(* IEC 61131-3 sources: SortJet_MasterSPS_Aufbau.fbsproj/07_Auftragsverwaltung/Auftragsspeicher, 3 files *)

(* ---- AuftragsSpeicher.fb.st ---- *)
(* METADATA
{
	"v3Meta": {
		"objectGuid": "f0eea758-4d67-47c3-84cf-9e26ec72588d"
	}
}
*)
FUNCTION_BLOCK AuftragsSpeicher
VAR_INPUT
  bpReset:BOOL;
  bpNeuerAuftrag:BOOL;
  bpNaechsterAuftrag :BOOL;
  NeuerAuftrag : Auftragsdaten_ST;
END_VAR
VAR_OUTPUT
  bpFehler:BOOL;
  bpAuftragverfuegbar:BOOL:=FALSE;
  AktAuftrag  :Auftragsdaten_ST;
END_VAR
VAR
  MerkerAuftrag :Auftragsdaten_ST;
END_VAR
(* Hinweis:
   - Auftragsdaten- Speicher fuer die " SHUTTLE "
*)
IF bpNeuerAuftrag THEN
  bpNeuerAuftrag:=FALSE;
  MerkerAuftrag := NeuerAuftrag;
  bpAuftragverfuegbar := TRUE;
END_IF

IF bpNaechsterAuftrag AND bpAuftragverfuegbar THEN
  bpNaechsterAuftrag := FALSE;
  AktAuftrag := MerkerAuftrag;
  bpAuftragverfuegbar:=FALSE;
END_IF

IF bpReset THEN
  bpFehler := FALSE;
  bpReset := FALSE;
  bpAuftragverfuegbar:=FALSE;
END_IF
END_FUNCTION_BLOCK

(* ---- Auftragsspeicher_FB.fb.st ---- *)
(* METADATA
{
	"v3Meta": {
		"objectGuid": "23ce62b1-5b0b-40f5-8f51-012d540e19cc"
	}
}
*)
FUNCTION_BLOCK Auftragsspeicher_FB
VAR_INPUT

  bpAktivieren     : BOOL := TRUE;
  bpWertAuslesen   : BOOL; // READ
  bpWerteSchreiben : BOOL; // WRITE
  bpReset          : BOOL; // RST

  // STRUCT
  stEingabeWert : Auftragsdaten_ST;

END_VAR
VAR_OUTPUT

  // BOOLEAN
  blWarteschlangeLeer : BOOL := TRUE;
  blWarteschlangeVoll : BOOL;

  // STRUCT
  stAusgabeWert  : Auftragsdaten_ST;

END_VAR
VAR

  // STRUCT
  warrlWarteSchlange : ARRAY[0..cINDEX] OF Auftragsdaten_ST;

  // INT
  ilReadPosition   : INT; // pr
  ilWritePosition  : INT; // pw
  iIndex           : INT;
END_VAR

VAR CONSTANT
  cINDEX : INT := 10;   // WICHTIG: Aenderungen an diesem Wert aendert die Anzahl der Elemente in der Warteschlange [FIFO]
END_VAR
//-------------------------------------------------------------------------------------------------
// BAUSTEIN: AUFTRAGSVERWALTUNG TRANSFERSHUTTLE
//-------------------------------------------------------------------------------------------------
IF ( bpReset ) THEN

  ilReadPosition      := 0;
  ilWritePosition     := 0;
  blWarteschlangeVoll := FALSE;
  blWarteschlangeLeer := TRUE;

  bpReset := FALSE;

ELSIF ( bpAktivieren ) THEN

  IF (  NOT blWarteschlangeLeer
       AND bpWertAuslesen )
  THEN
    stAusgabeWert := warrlWarteSchlange[ilReadPosition];
    ilReadPosition:= INCI(ilReadPosition, cINDEX );
    blWarteschlangeLeer := ( ilReadPosition = ilWritePosition );
    blWarteschlangeVoll := FALSE;
    bpWertAuslesen      := FALSE;
  END_IF;

  IF (  NOT blWarteschlangeVoll
       AND bpWerteSchreiben )
  THEN
    warrlWarteSchlange[ilWritePosition] := stEingabeWert;
    ilWritePosition := INCI( ilWritePosition, cINDEX );
    blWarteschlangeVoll := ( ilWritePosition = ilReadPosition );
    blWarteschlangeLeer := FALSE;
    bpWerteSchreiben    := FALSE;
  END_IF;

END_IF;
END_FUNCTION_BLOCK

(* ---- AuftragsSpeicherStationen.fb.st ---- *)
(* METADATA
{
	"v3Meta": {
		"objectGuid": "2fba16dc-56bd-4c56-9768-dbe33d4a7ec0"
	}
}
*)
FUNCTION_BLOCK AuftragsSpeicherStationen
VAR_INPUT

  // BOOLEAN
  bpReset            : BOOL;
  bpNeuerAuftrag     : BOOL;
  bpNaechsterAuftrag : BOOL;

  // STRUCT
  NeuerAuftrag : Auftragsdaten_ST;

END_VAR
VAR_OUTPUT

  // BOOLEAN
  bpFehler             : BOOL;
  bpAuftragverfuegbar : BOOL := FALSE;

  // STRUCT
  AktAuftrag : Auftragsdaten_ST;

END_VAR
VAR

  // STRUCT
  MerkerAuftrag :Auftragsdaten_ST;

END_VAR
(* Hinweis:
   - Auftragsdaten- Speicher fuer die " STATIONEN "
*)
IF ( bpNeuerAuftrag ) THEN
  bpNeuerAuftrag:=FALSE;
  MerkerAuftrag := NeuerAuftrag;
  bpAuftragverfuegbar := TRUE;
END_IF

IF ( bpNaechsterAuftrag AND bpAuftragverfuegbar ) THEN
  bpNaechsterAuftrag := FALSE;
  AktAuftrag := MerkerAuftrag;
  bpAuftragverfuegbar:=FALSE;
END_IF

IF ( bpReset ) THEN
  bpFehler := FALSE;
  bpReset := FALSE;
  bpAuftragverfuegbar:=FALSE;
END_IF
END_FUNCTION_BLOCK
